Fanuc KAREL source: kb00071.KL

-- PROVISIONAL review KL for V770-1; original PC SHA256 7c14a6db0779d05c4ad1e5ff25c4c2bfa06aeb584aef942bf280c9e918650768
-- Incomplete behavior may be omitted. Consult companion uncertainty JSON. Do not deploy.
PROGRAM KB00071
%NOLOCKGROUP
VAR
  P1 : REAL
  RESULT : REAL
BEGIN
  -- UNRESOLVED_PC offsets 5-16; opcodes 2E,23
  -- UNRESOLVED_PC offsets 21-36; opcodes 27,22,76,23
  -- UNRESOLVED_PC offsets 41-45; opcodes 7F
END KB00071
